(* IEC 61131-3 sources: guidance-for-physical-ai-production-designer-on-aws/source/plan2cell/crates/bt2plc/templates/codesys/device/DUT, 12 files *)

(* ---- E_PlayerState.st ---- *)
(*
 * E_PlayerState
 * States of FB_ProgramPlayer (robot side of the bt2plc zone protocol).
 * Device simulator {{ROBOT_TAG}} ({{ROBOT_NS}}), cell {{CELL_ID}}. Generated by {{GENERATOR}}.
 *)

TYPE E_PlayerState :
(
    PS_IDLE         := 0,    (* No program, pose held *)
    PS_NEXT_OP      := 10,   (* Advance to the next op: wStep := k, REQUEST := mask *)
    PS_WAIT_GRANT   := 20,   (* Wait (GRANT AND mask) = mask *)
    PS_DELAY        := 30,   (* Start delay of the op *)
    PS_MOVE         := 40,   (* Trajectory / blind home move *)
    PS_HOLD         := 50,   (* Hold at the end pose *)
    PS_WAIT_RELEASE := 60,   (* REQUEST := 0, wait (GRANT AND mask) = 0 *)
    PS_DONE         := 90,   (* Program finished *)
    PS_ERROR        := 99    (* Program aborted with an error *)
);
END_TYPE

(* ---- E_ProgramState.st ---- *)
(*
 * E_ProgramState
 * VW VASS standard - robot program states.
 * Device simulator {{ROBOT_TAG}} ({{ROBOT_NS}}), cell {{CELL_ID}}. Generated by {{GENERATOR}}.
 *)

TYPE E_ProgramState :
(
    PRG_IDLE     := 0,
    PRG_RUNNING  := 1,
    PRG_STOPPED  := 2,
    PRG_PAUSED   := 3,
    PRG_FINISHED := 4,
    PRG_ERROR    := 5
);
END_TYPE

(* ---- E_RobotMode.st ---- *)
(*
 * E_RobotMode
 * VW VASS standard - KUKA KR C4 robot operating modes.
 * Device simulator {{ROBOT_TAG}} ({{ROBOT_NS}}), cell {{CELL_ID}}. Generated by {{GENERATOR}}.
 *)

TYPE E_RobotMode :
(
    MODE_UNKNOWN := 0,
    MODE_T1      := 1,       (* Test mode 1 - reduced speed *)
    MODE_T2      := 2,       (* Test mode 2 - programmed speed *)
    MODE_AUT     := 3,       (* Automatic mode *)
    MODE_EXT     := 4        (* External automatic - PLC controlled *)
);
END_TYPE

(* ---- ST_OpDef.st ---- *)
(*
 * ST_OpDef
 * One op of the bt2plc robot program (row of GVL_Program.aOps).
 * Op k plays waypoints GVL_Program.aWp[nFirstWp..nLastWp] under the zone mask dwZoneMask.
 * Blind home op: bBlindHome = TRUE, nFirstWp = nLastWp = 0 (joint move to arHomeDeg over R_HOME_S).
 * Device simulator {{ROBOT_TAG}} ({{ROBOT_NS}}), cell {{CELL_ID}}. Generated by {{GENERATOR}}.
 *)

TYPE ST_OpDef :
STRUCT
    sName           : STRING(32);   (* Operation id, e.g. 'W01' *)
    nFirstWp        : INT;          (* First waypoint index in aWp (0 = none) *)
    nLastWp         : INT;          (* Last waypoint index in aWp (0 = none) *)
    dwZoneMask      : DWORD;        (* REQUEST/GRANT bits (zones 0..30, bit 31 = permit) *)
    tDelay          : TIME;         (* Start delay after the grant *)
    tHold           : TIME;         (* Hold time at the end pose *)
    rDelay_s        : REAL;         (* Start delay in s (used by FB_ProgramPlayer) *)
    rHold_s         : REAL;         (* Hold time in s (used by FB_ProgramPlayer) *)
    rVelScale       : REAL;         (* Velocity scale of the trajectory (1.0 = nominal) *)
    bBlindHome      : BOOL;         (* TRUE = blind joint move to the home pose *)
END_STRUCT
END_TYPE

(* ---- ST_PROFIsafe_Trailer.st ---- *)
(*
 * ST_PROFIsafe_Trailer
 * PROFIsafe trailer - 4 bytes appended by the safety layer (status + 3-byte CRC).
 * Device simulator {{ROBOT_TAG}} ({{ROBOT_NS}}), cell {{CELL_ID}}. Generated by {{GENERATOR}}.
 *)

TYPE ST_PROFIsafe_Trailer :
STRUCT
    byStatus        : BYTE;                     (* Status/Control byte *)
    abyCRC          : ARRAY[0..2] OF BYTE;      (* 3-byte CRC *)
END_STRUCT
END_TYPE

(* ---- ST_SafeInput.st ---- *)
(*
 * ST_SafeInput
 * PROFIsafe (Slot 1 - FDIO64) safe inputs: robot -> PLC, 8 bytes user data.
 * GSDML: 8x Unsigned8 Input + F_MessageTrailer4Byte.
 * Device simulator {{ROBOT_TAG}} ({{ROBOT_NS}}), cell {{CELL_ID}}. Generated by {{GENERATOR}}.
 *)

TYPE ST_SafeInput :
STRUCT
    (* Byte 0: Safe robot status *)
    bSafe_DrivesOK          : BOOL;   (* Bit 0: Safe drives monitoring OK *)
    bSafe_RobotStopped      : BOOL;   (* Bit 1: Robot safely stopped (SOS/SS1) *)
    bSafe_ReducedSpeed      : BOOL;   (* Bit 2: Safe reduced speed active (SLS) *)
    bSafe_AxisMonitoring    : BOOL;   (* Bit 3: Safe axis range monitoring OK *)
    bSafe_ToolOK            : BOOL;   (* Bit 4: Safe tool monitoring OK *)
    bSafe_WorkspaceOK       : BOOL;   (* Bit 5: Safe workspace monitoring OK *)
    bSafe_Reserved06        : BOOL;   (* Bit 6: Reserved *)
    bSafe_Reserved07        : BOOL;   (* Bit 7: Reserved *)

    (* Byte 1: Safe gate/zone status *)
    bSafe_Gate1Closed       : BOOL;   (* Bit 0: Safety gate 1 closed *)
    bSafe_Gate2Closed       : BOOL;   (* Bit 1: Safety gate 2 closed *)
    bSafe_Gate3Closed       : BOOL;   (* Bit 2: Safety gate 3 closed *)
    bSafe_LightCurtainOK    : BOOL;   (* Bit 3: Light curtain free *)
    bSafe_EStopOK           : BOOL;   (* Bit 4: E-Stop not pressed (NC) *)
    bSafe_EnablingDevice    : BOOL;   (* Bit 5: Enabling device pressed (T1/T2) *)
    bSafe_OperatorSafe      : BOOL;   (* Bit 6: Operator protection OK *)
    bSafe_Reserved17        : BOOL;   (* Bit 7: Reserved *)

    (* Byte 2: Extended safe status *)
    bSafe_STO_Active        : BOOL;   (* Bit 0: Safe Torque Off active *)
    bSafe_SS1_Active        : BOOL;   (* Bit 1: Safe Stop 1 active *)
    bSafe_SS2_Active        : BOOL;   (* Bit 2: Safe Stop 2 active *)
    bSafe_SOS_Active        : BOOL;   (* Bit 3: Safe Operating Stop active *)
    bSafe_SLS_Active        : BOOL;   (* Bit 4: Safely-Limited Speed active *)
    bSafe_SLP_Active        : BOOL;   (* Bit 5: Safely-Limited Position active *)
    bSafe_Reserved26        : BOOL;   (* Bit 6: Reserved *)
    bSafe_FaultPresent      : BOOL;   (* Bit 7: Safety fault present *)

    (* Bytes 3-7: Additional safe signals *)
    bySafe_UserInput3       : BYTE;   (* Byte 3: User safe input *)
    bySafe_UserInput4       : BYTE;   (* Byte 4: User safe input *)
    bySafe_UserInput5       : BYTE;   (* Byte 5: User safe input *)
    bySafe_UserInput6       : BYTE;   (* Byte 6: User safe input *)
    bySafe_UserInput7       : BYTE;   (* Byte 7: User safe input *)
END_STRUCT
END_TYPE

(* ---- ST_SafeOutput.st ---- *)
(*
 * ST_SafeOutput
 * PROFIsafe (Slot 1 - FDIO64) safe outputs: PLC -> robot, 8 bytes user data.
 * GSDML: 8x Unsigned8 Output + F_MessageTrailer4Byte.
 * Device simulator {{ROBOT_TAG}} ({{ROBOT_NS}}), cell {{CELL_ID}}. Generated by {{GENERATOR}}.
 *)

TYPE ST_SafeOutput :
STRUCT
    (* Byte 0: Safe control from PLC *)
    bSafe_DriveEnable       : BOOL;   (* Bit 0: Enable drives (safe channel) *)
    bSafe_ExternalEStop     : BOOL;   (* Bit 1: External E-Stop request *)
    bSafe_SafeStop1         : BOOL;   (* Bit 2: Request Safe Stop 1 *)
    bSafe_SafeStop2         : BOOL;   (* Bit 3: Request Safe Stop 2 *)
    bSafe_ReducedSpeedReq   : BOOL;   (* Bit 4: Request safe reduced speed *)
    bSafe_GateOverride      : BOOL;   (* Bit 5: Gate override (maintenance) *)
    bSafe_Reserved06        : BOOL;   (* Bit 6: Reserved *)
    bSafe_Reserved07        : BOOL;   (* Bit 7: Reserved *)

    (* Byte 1: Safe zone control *)
    bSafe_Zone1Enable       : BOOL;   (* Bit 0: Enable workspace zone 1 *)
    bSafe_Zone2Enable       : BOOL;   (* Bit 1: Enable workspace zone 2 *)
    bSafe_Zone3Enable       : BOOL;   (* Bit 2: Enable workspace zone 3 *)
    bSafe_Zone4Enable       : BOOL;   (* Bit 3: Enable workspace zone 4 *)
    bSafe_Reserved14        : BOOL;   (* Bit 4: Reserved *)
    bSafe_Reserved15        : BOOL;   (* Bit 5: Reserved *)
    bSafe_Reserved16        : BOOL;   (* Bit 6: Reserved *)
    bSafe_Reserved17        : BOOL;   (* Bit 7: Reserved *)

    (* Bytes 2-7: Additional safe control *)
    bySafe_UserOutput2      : BYTE;   (* Byte 2: User safe output *)
    bySafe_UserOutput3      : BYTE;   (* Byte 3: User safe output *)
    bySafe_UserOutput4      : BYTE;   (* Byte 4: User safe output *)
    bySafe_UserOutput5      : BYTE;   (* Byte 5: User safe output *)
    bySafe_UserOutput6      : BYTE;   (* Byte 6: User safe output *)
    bySafe_UserOutput7      : BYTE;   (* Byte 7: User safe output *)
END_STRUCT
END_TYPE

(* ---- ST_VASS_ControlWord.st ---- *)
(*
 * ST_VASS_ControlWord
 * VASS PLC control word - output bytes 0-1 (PLC -> robot), Slot 2 DIO256.
 * Device simulator {{ROBOT_TAG}} ({{ROBOT_NS}}), cell {{CELL_ID}}. Generated by {{GENERATOR}}.
 *)

TYPE ST_VASS_ControlWord :
STRUCT
    (* Byte 0 *)
    bDrivesOn           : BOOL;   (* Bit 0: Enable drives *)
    bProgStart          : BOOL;   (* Bit 1: Start program *)
    bProgStop           : BOOL;   (* Bit 2: Stop program *)
    bProgCancel         : BOOL;   (* Bit 3: Cancel program *)
    bModeRequest        : BOOL;   (* Bit 4: Request EXT mode *)
    bReset              : BOOL;   (* Bit 5: Reset error *)
    bHomeRequest        : BOOL;   (* Bit 6: Move to home *)
    bConfirm            : BOOL;   (* Bit 7: Confirm/acknowledge *)

    (* Byte 1 *)
    bJobRequest         : BOOL;   (* Bit 8: New job request *)
    bGripperOpen        : BOOL;   (* Bit 9: Open gripper *)
    bGripperClose       : BOOL;   (* Bit 10: Close gripper *)
    bPeriphRelease      : BOOL;   (* Bit 11: Release peripheral *)
    bSpeedOverride      : BOOL;   (* Bit 12: Apply speed override *)
    bReserved13         : BOOL;   (* Bit 13: Reserved *)
    bReserved14         : BOOL;   (* Bit 14: Reserved *)
    bReserved15         : BOOL;   (* Bit 15: Reserved *)
END_STRUCT
END_TYPE

(* ---- ST_VASS_InputTelegram.st ---- *)
(*
 * ST_VASS_InputTelegram
 * Full VASS input telegram - 32 bytes (robot -> PLC), Slot 2 DIO256 inputs.
 * bt2plc use: bytes 4-5 wCurrentStep = op index (GVL_Program.STEP_BYTE),
 *             bytes 16-27 joint angles A1..A6 (FB_JointAngleEncoder),
 *             bytes 28-31 zone REQUEST DWORD LE (GVL_Program.REQ_BYTE).
 * Device simulator {{ROBOT_TAG}} ({{ROBOT_NS}}), cell {{CELL_ID}}. Generated by {{GENERATOR}}.
 *)

TYPE ST_VASS_InputTelegram :
STRUCT
    stStatusWord        : ST_VASS_StatusWord;     (* Bytes 0-1:   Status word *)
    wActiveJobNr        : WORD;                   (* Bytes 2-3:   Active job number *)
    wCurrentStep        : WORD;                   (* Bytes 4-5:   Current program step *)
    wSpeedActual        : WORD;                   (* Bytes 6-7:   Actual speed % *)
    wActiveToolNr       : WORD;                   (* Bytes 8-9:   Active tool number *)
    wErrorCode          : WORD;                   (* Bytes 10-11: Active error code *)
    wWarningCode        : WORD;                   (* Bytes 12-13: Active warning code *)
    wPositionX          : INT;                    (* Bytes 14-15: Position X (0.1mm) *)
    wPositionY          : INT;                    (* Bytes 16-17: Position Y (0.1mm) *)
    wPositionZ          : INT;                    (* Bytes 18-19: Position Z (0.1mm) *)
    wUserWord10         : WORD;                   (* Bytes 20-21: User data *)
    wUserWord11         : WORD;                   (* Bytes 22-23: User data *)
    wUserWord12         : WORD;                   (* Bytes 24-25: User data *)
    wUserWord13         : WORD;                   (* Bytes 26-27: User data *)
    wUserWord14         : WORD;                   (* Bytes 28-29: User data *)
    wUserWord15         : WORD;                   (* Bytes 30-31: User data *)
END_STRUCT
END_TYPE

(* ---- ST_VASS_OutputTelegram.st ---- *)
(*
 * ST_VASS_OutputTelegram
 * Full VASS output telegram - 32 bytes (PLC -> robot), Slot 2 DIO256 outputs.
 * bt2plc use: bytes 4-5 PLAN_ID WORD LE during a production job (GVL_Program.PLAN_ID_BYTE),
 *             bytes 12-15 zone GRANT DWORD LE (GVL_Program.GRANT_BYTE).
 * Device simulator {{ROBOT_TAG}} ({{ROBOT_NS}}), cell {{CELL_ID}}. Generated by {{GENERATOR}}.
 *)

TYPE ST_VASS_OutputTelegram :
STRUCT
    stControlWord       : ST_VASS_ControlWord;    (* Bytes 0-1:   Control word *)
    wJobNr              : WORD;                   (* Bytes 2-3:   Requested job number *)
    wParameter1         : WORD;                   (* Bytes 4-5:   Parameter 1 *)
    wParameter2         : WORD;                   (* Bytes 6-7:   Parameter 2 *)
    wSpeedOverride      : WORD;                   (* Bytes 8-9:   Speed override % *)
    wToolRequest        : WORD;                   (* Bytes 10-11: Tool change request *)
    wUserWord6          : WORD;                   (* Bytes 12-13: User command data *)
    wUserWord7          : WORD;                   (* Bytes 14-15: User command data *)
    wUserWord8          : WORD;                   (* Bytes 16-17: User command data *)
    wUserWord9          : WORD;                   (* Bytes 18-19: User command data *)
    wUserWord10         : WORD;                   (* Bytes 20-21: User command data *)
    wUserWord11         : WORD;                   (* Bytes 22-23: User command data *)
    wUserWord12         : WORD;                   (* Bytes 24-25: User command data *)
    wUserWord13         : WORD;                   (* Bytes 26-27: User command data *)
    wUserWord14         : WORD;                   (* Bytes 28-29: User command data *)
    wUserWord15         : WORD;                   (* Bytes 30-31: User command data *)
END_STRUCT
END_TYPE

(* ---- ST_VASS_StatusWord.st ---- *)
(*
 * ST_VASS_StatusWord
 * VASS robot status word - input bytes 0-1 (robot -> PLC), Slot 2 DIO256.
 * Device simulator {{ROBOT_TAG}} ({{ROBOT_NS}}), cell {{CELL_ID}}. Generated by {{GENERATOR}}.
 *)

TYPE ST_VASS_StatusWord :
STRUCT
    (* Byte 0 *)
    bDrivesPowered      : BOOL;   (* Bit 0: Drives are powered on *)
    bProgRunning        : BOOL;   (* Bit 1: Program is running *)
    bAtHome             : BOOL;   (* Bit 2: Robot at home position *)
    bInPosition         : BOOL;   (* Bit 3: Robot in target position *)
    bModeExt            : BOOL;   (* Bit 4: External automatic mode active *)
    bReady              : BOOL;   (* Bit 5: Robot ready for command *)
    bError              : BOOL;   (* Bit 6: Error present *)
    bWarning            : BOOL;   (* Bit 7: Warning present *)

    (* Byte 1 *)
    bSafetyGateOK       : BOOL;   (* Bit 8: Safety gate closed *)
    bEStopNotActive     : BOOL;   (* Bit 9: E-Stop NOT active (NC logic) *)
    bProgFinished       : BOOL;   (* Bit 10: Program/job finished *)
    bJobAcknowledge     : BOOL;   (* Bit 11: Job number acknowledged *)
    bToolActive         : BOOL;   (* Bit 12: Tool/gripper active *)
    bPartPresent        : BOOL;   (* Bit 13: Part present in gripper *)
    bPeriphReady        : BOOL;   (* Bit 14: Peripheral devices ready *)
    bMaintRequired      : BOOL;   (* Bit 15: Maintenance required *)
END_STRUCT
END_TYPE

(* ---- ST_Waypoint.st ---- *)
(*
 * ST_Waypoint
 * One trajectory waypoint (row of GVL_Program.aWp). Flat fields for portability.
 * rT = seconds from op start; angles in degrees (KUKA A1..A6 after joint sign/offset mapping).
 * Device simulator {{ROBOT_TAG}} ({{ROBOT_NS}}), cell {{CELL_ID}}. Generated by {{GENERATOR}}.
 *)

TYPE ST_Waypoint :
STRUCT
    rT              : REAL;         (* Time from op start (s) *)
    rA1             : REAL;         (* Axis 1 (deg) *)
    rA2             : REAL;         (* Axis 2 (deg) *)
    rA3             : REAL;         (* Axis 3 (deg) *)
    rA4             : REAL;         (* Axis 4 (deg) *)
    rA5             : REAL;         (* Axis 5 (deg) *)
    rA6             : REAL;         (* Axis 6 (deg) *)
END_STRUCT
END_TYPE
